(* PLC project forms.project, CODESYS CODESYS V3.5 SP17 Patch 3 *)
(* stored: creationDateTime 2026-10-20T03:44:11.3196869, modificationDateTime 1601-01-01T03:00:00 *)

TYPE ST_Probe : STRUCT
  a : INT;
  b : BOOL;
END_STRUCT;
END_TYPE

FUNCTION_BLOCK FB_ProbeOop
  VAR_INPUT
    xIn : BOOL;
  END_VAR
  VAR
    iState : INT;
  END_VAR

                  iState := iState + 1;

                

ACTION ActClear:
                      iState := 0;

                    
END_ACTION

METHOD Reset : BOOL
  VAR_INPUT
    iTo : INT;
  END_VAR
                        iState := iTo;
Reset := TRUE;

                      
END_METHOD

PROPERTY State : INT
GET
                          State := iState;

                        
END_GET
SET
                          iState := State;

                        
END_SET
END_PROPERTY
END_FUNCTION_BLOCK

PROGRAM PRG_ProbeMain
  VAR
    fbOop : FB_ProbeOop;
  END_VAR

                  fbOop(xIn := GVL_Probe.xFlag);
GVL_Probe.diHours := GVL_Probe.diHours + 1;

                
END_PROGRAM

CONFIGURATION Application
  RESOURCE Application ON PLC
    {attribute 'qualified_only'}
    VAR_GLOBAL  (* GVL_Probe *)
      xFlag : BOOL;
      iCount : INT := 5;
      rTotal : REAL;
      diHours : DINT;
    END_VAR
    TASK Task_Fast(INTERVAL := T#10ms, PRIORITY := 1);
    TASK Task_Free(PRIORITY := 20);
    PROGRAM PRG_ProbeMain WITH Task_Fast : PRG_ProbeMain;
  END_RESOURCE
END_CONFIGURATION
